// TIA Portal project "SortingStation" (V19)

(* hardware
DEVICE "S7-1500/ET200MP station_1"  S7-1500 station
   slot 0: "Rail_0"  Rack  6ES7 590-1***0-0AA0
   slot 1: "PLC_1"  CPU 1511-1 PN  6ES7 511-1AK02-0AB0  V2.9
      slot 3: "CPU display_1"  6ES7591-1AA00-0AA0
      slot 32768: "PROFINET interface_1"  X1
         slot 32769: "Port_1"  X1 P1
         slot 32770: "Port_2"  X1 P2
      slot 34817: "Virtual CP interface port_1"  Virtual CP interface port  Virtual CP interface port
   slot 2: "DI 16x24VDC BA_1"  DI 16x24VDC BA  6ES7 521-1BH10-0AA0  V1.1
   slot 3: "DQ 16x24VDC/0.5A BA_1"  DQ 16x24VDC/0.5A BA  6ES7 522-1BH10-0AA0  V1.1
   slot 4: "AI 4xU/I/RTD/TC ST_1"  AI 4xU/I/RTD/TC ST  6ES7 531-7QD00-0AB0  V1.0
DEVICE "HMI_1"  TP700 Comfort
   slot 0: "HMI_1"  TP700 Comfort  6AV2 124-0GC01-0AX0  17.0.0.0
   slot 1: "HMI_RT_1"  TP700 Comfort  6AV2 124-0GC01-0AX0  17.0.0.0
   slot 5: "HMI_1.IE_CP_1"  PROFINET Interface  17.0.0.0
      slot 1: "PROFINET Interface_1"  PROFINET Interface
         slot 1: "Port_1"  Port
         slot 2: "Port_2"  Port
   slot 7: "HMI_1.MPI/DP_CP_1"  MPI/DP Interface  17.0.0.0
*)

// ===== PLC "PLC_1"  CPU 1511-1 PN =====

VAR_GLOBAL   // PLC tag table "Default tag table"
   "System_Byte" AT %MB1 : Byte;
   "FirstScan" AT %M1.0 : Bool;
   "DiagStatusUpdate" AT %M1.1 : Bool;
   "AlwaysTRUE" AT %M1.2 : Bool;
   "AlwaysFALSE" AT %M1.3 : Bool;
   "Clock_Byte" AT %MB0 : Byte;
   "Clock_10Hz" AT %M0.0 : Bool;
   "Clock_5Hz" AT %M0.1 : Bool;
   "Clock_2.5Hz" AT %M0.2 : Bool;
   "Clock_2Hz" AT %M0.3 : Bool;
   "Clock_1.25Hz" AT %M0.4 : Bool;
   "Clock_1Hz" AT %M0.5 : Bool;
   "Clock_0.625Hz" AT %M0.6 : Bool;
   "Clock_0.5Hz" AT %M0.7 : Bool;
END_VAR

VAR_GLOBAL   // PLC tag table "IO_Tags"
   "PB_Start" AT %I0.0 : Bool;   // Start pushbutton, NO contact
   "PB_Stop" AT %I0.1 : Bool;   // Stop pushbutton, NC contact
   "PB_Reset" AT %I0.2 : Bool;   // Alarm reset pushbutton
   "ESTOP_OK" AT %I0.3 : Bool;   // Emergency stop circuit, 1 = healthy
   "S_Entry" AT %I0.4 : Bool;   // Part entry sensor
   "S_Defective" AT %I0.5 : Bool;   // Defective part signal
   "Motor_Overload_OK" AT %I0.6 : Bool;   // Motor overload relay, NC, 1 = healthy
   "AI_MotorTemp" AT %IW64 : Int;   // Motor temperature, raw analog value 0..27648
   "K_Motor" AT %Q0.0 : Bool;   // Conveyor motor contactor
   "L_Run" AT %Q0.1 : Bool;   // Green lamp, running
   "L_Fault" AT %Q0.2 : Bool;   // Red lamp, fault
   "L_Idle" AT %Q0.3 : Bool;   // Yellow lamp, idle
   "Y_Diverter" AT %Q0.4 : Bool;   // Diverter actuator for rejected parts
   "Horn" AT %Q0.5 : Bool;   // Alarm horn
END_VAR

TYPE "udt_Station"
   STRUCT
      State : Int;   // 0=Idle, 1=Running, 2=Fault
      FaultCode : Word := 0;   // bit0=EStop, bit1=Overload, bit2=OverTemp, bit3=Jam
      CntGood : DInt := 0;   // Count of good parts
      CntReject : DInt;   // Count of rejected parts
      MotorTemp : Real;   // Scaled motor temperature in degC
      TempLimit : Real := 80.0;   // Max allowed motor temperature in degC
      HMI_Start : Bool;   // Start command from HMI
      HMI_Stop : Bool;   // Stop command from HMI
      HMI_Reset : Bool;   // Alarm reset command from HMI
      HMI_ResetCnt : Bool;   // Counter reset command from HMI
   END_STRUCT;
END_TYPE

DATA_BLOCK "DB_Station"   // DB1
{ S7_Optimized_Access := 'TRUE' }
VERSION : 0.1
BEGIN
END_DATA_BLOCK

DATA_BLOCK "iDB_Station"   // DB2
{ S7_Optimized_Access := 'TRUE' }
VERSION : 0.1
// stored: InstanceOfName FB_Station
"FB_Station"
BEGIN
END_DATA_BLOCK

FUNCTION_BLOCK "FB_Motor"   // FB1, LAD
{ S7_Optimized_Access := 'TRUE' }
VERSION : 0.1
   VAR_INPUT
      Start : Bool;   // Start command, 1 = start requested
      Stop : Bool;   // Stop command, 1 = stop requested
      Permissive : Bool;   // Interlock, 1 = all conditions healthy
   END_VAR
   VAR_OUTPUT
      Run : Bool;   // Motor run command
   END_VAR
   VAR
      RunMem : Bool;   // Seal-in memory bit
   END_VAR
BEGIN

REGION Network 1: Seal-in memory bit
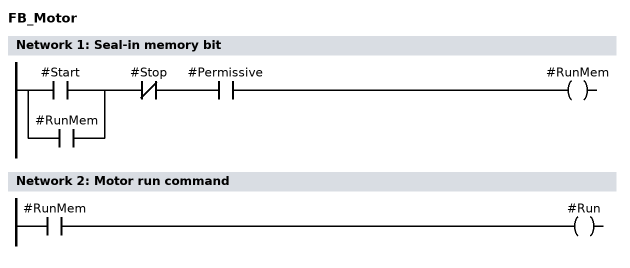
   RUNG wire#powerrail
      Contact( #Start )
      wire#w1
      I_Contact( #Stop )
      Contact( #Permissive )
      Coil( #RunMem )
   END_RUNG
   RUNG wire#powerrail
      Contact( #RunMem )
   END_RUNG wire#w1
   // the same network as SCL:
   #RunMem := (#Start OR #RunMem) AND NOT #Stop AND #Permissive;
END_REGION

REGION Network 2: Motor run command
   RUNG wire#powerrail
      Contact( #RunMem )
      Coil( #Run )
   END_RUNG
   // the same network as SCL:
   #Run := #RunMem;
END_REGION
END_FUNCTION_BLOCK

FUNCTION_BLOCK "FB_Station"   // FB2, SCL
{ S7_Optimized_Access := 'TRUE' }
VERSION : 0.1
   VAR_INPUT
      PB_Start : Bool;   // Start pushbutton, NO
      PB_Stop : Bool;   // Stop pushbutton, NC, 0 = pressed
      PB_Reset : Bool;   // Alarm reset pushbutton
      ESTOP_OK : Bool;   // Emergency stop circuit, 1 = healthy
      S_Entry : Bool;   // Part entry sensor
      S_Defective : Bool;   // Defective part signal
      Motor_Overload_OK : Bool;   // Overload relay, 1 = healthy
      Clock1Hz : Bool;   // 1 Hz clock bit for blinking
   END_VAR
   VAR_OUTPUT
      K_Motor : Bool;   // Conveyor motor contactor
      L_Run : Bool;   // Green lamp
      L_Fault : Bool;   // Red lamp, blinking
      L_Idle : Bool;   // Yellow lamp
      Y_Diverter : Bool;   // Diverter for rejected parts
      Horn : Bool;   // Alarm horn
   END_VAR
   VAR_IN_OUT
      Station : "udt_Station";   // Station data, passed from DB_Station
   END_VAR
   VAR
      motor : "FB_Motor";   // Motor control instance
      tonJam : TON_TIME;   // Jam detection timer
      tpDiverter : TP_TIME;   // Diverter pulse timer
   END_VAR
   VAR RETAIN
      ctuGood : CTU_DINT;   // Good parts counter
      ctuReject : CTU_DINT;   // Rejected parts counter
   END_VAR
   VAR
      rtStart : R_TRIG;   // Start edge
      rtReset : R_TRIG;   // Reset edge
      rtEntry : R_TRIG;   // Entry sensor edge
   END_VAR
   VAR_TEMP
      stopCmd : Bool;
      anyFault : Bool;
      fEStop : Bool;
      fOverload : Bool;
      fOverTemp : Bool;
      fJam : Bool;
      goodPulse : Bool;
      rejectPulse : Bool;
   END_VAR
BEGIN
   // =====================================================
   // FB_Station : sorting station main logic
   // States: 0 = Idle, 1 = Running, 2 = Fault
   // FaultCode: bit0 EStop, bit1 Overload, bit2 OverTemp, bit3 Jam
   // =====================================================

   // ---- 1. Edge detection and commands ----
   #rtStart(CLK := #PB_Start OR #Station.HMI_Start);
   #rtReset(CLK := #PB_Reset OR #Station.HMI_Reset);
   #rtEntry(CLK := #S_Entry);

   // PB_Stop is NC: 0 = pressed
   #stopCmd := (NOT #PB_Stop) OR #Station.HMI_Stop;

   // ---- 2. Fault detection (live conditions) ----
   #fEStop := NOT #ESTOP_OK;
   #fOverload := NOT #Motor_Overload_OK;
   #fOverTemp := #Station.MotorTemp > #Station.TempLimit;

   // Jam: entry sensor active longer than 5 s while running
   #tonJam(IN := #S_Entry AND (#Station.State = 1),
           PT := T#5s);
   #fJam := #tonJam.Q;

   #anyFault := #fEStop OR #fOverload OR #fOverTemp OR #fJam;

   // ---- 3. Latched fault code ----
   // Reset clears the code first, then active faults set their bits again
   IF #rtReset.Q THEN
       #Station.FaultCode := W#16#0000;
   END_IF;

   IF #fEStop THEN
       #Station.FaultCode := #Station.FaultCode OR W#16#0001;
   END_IF;
   IF #fOverload THEN
       #Station.FaultCode := #Station.FaultCode OR W#16#0002;
   END_IF;
   IF #fOverTemp THEN
       #Station.FaultCode := #Station.FaultCode OR W#16#0004;
   END_IF;
   IF #fJam THEN
       #Station.FaultCode := #Station.FaultCode OR W#16#0008;
   END_IF;

   // ---- 4. State machine ----
   CASE #Station.State OF
       0:  // Idle
           IF #anyFault THEN
               #Station.State := 2;
           ELSIF #rtStart.Q AND NOT #stopCmd THEN
               #Station.State := 1;
           END_IF;

       1:  // Running
           IF #anyFault THEN
               #Station.State := 2;
           ELSIF #stopCmd THEN
               #Station.State := 0;
           END_IF;

       2:  // Fault: leave only on reset with all faults cleared
           IF #rtReset.Q AND NOT #anyFault THEN
               #Station.State := 0;
           END_IF;

       ELSE
           #Station.State := 2;
   END_CASE;

   // ---- 5. Sorting logic (only while running) ----
   #goodPulse := FALSE;
   #rejectPulse := FALSE;

   IF (#Station.State = 1) AND #rtEntry.Q THEN
       IF #S_Defective THEN
           #rejectPulse := TRUE;
       ELSE
           #goodPulse := TRUE;
       END_IF;
   END_IF;

   #ctuGood(CU := #goodPulse,
            R := #Station.HMI_ResetCnt,
            PV := 99999999);
   #ctuReject(CU := #rejectPulse,
              R := #Station.HMI_ResetCnt,
              PV := 99999999);
   #Station.CntGood := #ctuGood.CV;
   #Station.CntReject := #ctuReject.CV;

   // Diverter: 2 s pulse for each rejected part
   #tpDiverter(IN := #rejectPulse,
               PT := T#2s);
   #Y_Diverter := #tpDiverter.Q AND (#Station.State = 1);

   // ---- 6. Motor control ----
   // Permissive drops the motor in Idle and Fault
   #motor(Start := #PB_Start OR #Station.HMI_Start,
          Stop := #stopCmd,
          Permissive := (#Station.State = 1));
   #K_Motor := #motor.Run;

   // ---- 7. Lamps and horn ----
   #L_Idle := (#Station.State = 0);
   #L_Run := (#Station.State = 1);
   #L_Fault := (#Station.State = 2) AND #Clock1Hz;
   #Horn := (#Station.State = 2);
END_FUNCTION_BLOCK

ORGANIZATION_BLOCK "Main"   // OB1, LAD, ProgramCycle
TITLE = "Main Program Sweep (Cycle)"
{ S7_Optimized_Access := 'TRUE' }
VERSION : 0.1
   VAR_INPUT
      Initial_Call : Bool;   // Initial call of this OB
      Remanence : Bool;   // =True, if remanent data are available
   END_VAR
   VAR_TEMP
      normTemp : Real;   // Normalized temperature 0.0 to 1.0
   END_VAR
BEGIN

REGION Network 1
   // Scale raw analog value 0..27648 to 0..150 degC
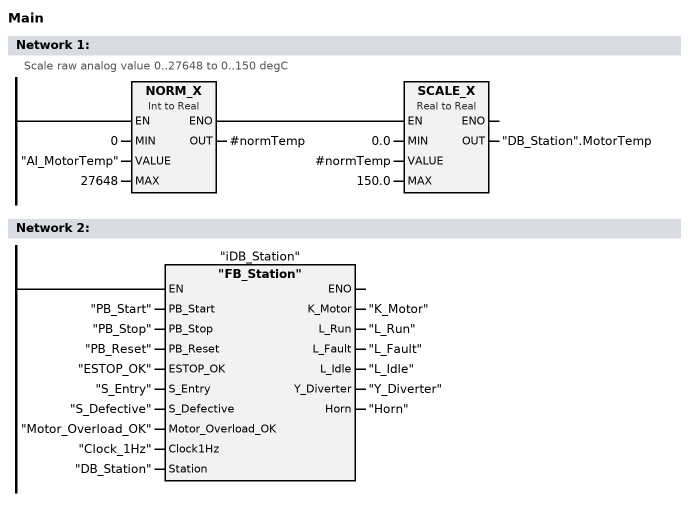
   RUNG wire#powerrail
      { S7_Templates := "[SrcType := Int, DestType := Real]" } Normalize(min := 0, value := "AI_MotorTemp", max := 27648, out => #normTemp)
      { S7_Templates := "[SrcType := Real, DestType := Real]" } Scale(min := 0.0, value := #normTemp, max := 150.0, out => "DB_Station".MotorTemp)
   END_RUNG
   // the same network as SCL:
   #normTemp := NORM_X(MIN := 0, VALUE := "AI_MotorTemp", MAX := 27648);
   "DB_Station".MotorTemp := SCALE_X(MIN := 0.0, VALUE := #normTemp, MAX := 150.0);
END_REGION

REGION Network 2
   RUNG wire#powerrail
      "iDB_Station"(PB_Start := "PB_Start", PB_Stop := "PB_Stop", PB_Reset := "PB_Reset", ESTOP_OK := "ESTOP_OK", S_Entry := "S_Entry", S_Defective := "S_Defective", Motor_Overload_OK := "Motor_Overload_OK", Clock1Hz := "Clock_1Hz", Station := "DB_Station", K_Motor => "K_Motor", L_Run => "L_Run", L_Fault => "L_Fault", L_Idle => "L_Idle", Y_Diverter => "Y_Diverter", Horn => "Horn")
   END_RUNG
   // the same network as SCL:
   "iDB_Station"(PB_Start := "PB_Start",   // "FB_Station"
                 PB_Stop := "PB_Stop",
                 PB_Reset := "PB_Reset",
                 ESTOP_OK := "ESTOP_OK",
                 S_Entry := "S_Entry",
                 S_Defective := "S_Defective",
                 Motor_Overload_OK := "Motor_Overload_OK",
                 Clock1Hz := "Clock_1Hz",
                 Station := "DB_Station",
                 K_Motor => "K_Motor",
                 L_Run => "L_Run",
                 L_Fault => "L_Fault",
                 L_Idle => "L_Idle",
                 Y_Diverter => "Y_Diverter",
                 Horn => "Horn");
END_REGION
END_ORGANIZATION_BLOCK

ORGANIZATION_BLOCK "Startup"   // OB100, SCL, Startup
TITLE = "Complete Restart"
{ S7_Optimized_Access := 'TRUE' }
VERSION : 0.1
   VAR_INPUT
      LostRetentive : Bool;   // True if retentive data are lost
      LostRTC : Bool;   // True if date and time are lost
   END_VAR
BEGIN
   // =====================================================
   // OB100 Startup : runs once at every STOP to RUN transition
   // Puts the station in a known safe state
   // =====================================================
   "DB_Station".State := 0;
   "DB_Station".FaultCode := W#16#0000;

   "DB_Station".HMI_Start := FALSE;
   "DB_Station".HMI_Stop := FALSE;
   "DB_Station".HMI_Reset := FALSE;
   "DB_Station".HMI_ResetCnt := FALSE;
END_ORGANIZATION_BLOCK

(* ===== HMI "HMI_RT_1" =====
system functions are stored by id; their names below are inferred from use
connection "HMI_Connection_1": ETHERNET, S7_1500_OMS

HMI tags "Default tag table"
   "Tag_ScreenNumber" : UInt, internal
   "Station_State" : Int = PLC DB_Station.State, 1 s
   "Station_FaultCode" : Word = PLC DB_Station.FaultCode AT %DB1.DBW0, 1 s
   "Station_CntGood" : DInt = PLC DB_Station.CntGood AT %DB1.DBW0, 1 s
   "Station_CntReject" : DInt = PLC DB_Station.CntReject AT %DB1.DBD0, 1 s
   "Station_MotorTemp" : Real = PLC DB_Station.MotorTemp AT %DB1.DBD0, 1 s
   "Station_TempLimit" : Real = PLC DB_Station.TempLimit AT %DB1.DBD0, 1 s
   "Station_HMI_Start" : Bool = PLC DB_Station.HMI_Start AT %DB1.DBD0, 1 s
   "Station_HMI_Stop" : Bool = PLC DB_Station.HMI_Stop AT %DB1.DBX0.0, 1 s
   "Station_HMI_Reset" : Bool = PLC DB_Station.HMI_Reset AT %DB1.DBX0.0, 1 s
   "Station_HMI_ResetCnt" : Bool = PLC DB_Station.HMI_ResetCnt AT %DB1.DBX0.0, 1 s

screen "Root screen" 800x420, template "Template_1"
   on GenerateScreen: SetTag("Tag_ScreenNumber", 1)
   TextField "HmiScreenItemData" at 78,377 size 640x25; Text 'Welcome to HMI_1 (TP700 Comfort)!'
   TextField "Text field_1" at 31,11 size 209x34; Text 'Sorting Station'
   TextField "Text field_2" at 78,70 size 54x23; Text 'State'
   TextField "Text field_3" at 77,113 size 51x23; Text 'Good'
   TextField "Text field_4" at 54,157 size 86x23; Text 'Rejected'
   TextField "Text field_5" at 19,201 size 123x23; Text 'Temperature'
   TextField "Text field_6" at 43,247 size 99x23; Text 'Fault code'
   IOField "I/O field_1" at 142,67 size 96x32; FormatPattern 9
      ProcessValue <- "Station_State"
   IOField "I/O field_2" at 142,108 size 96x32; FormatPattern 99999
      ProcessValue <- "Station_CntGood"
   IOField "I/O field_3" at 143,152 size 96x32; FormatPattern 99999
      ProcessValue <- "Station_CntReject"
   IOField "I/O field_4" at 143,197 size 96x32; FormatPattern 999.9
      ProcessValue <- "Station_MotorTemp"
   IOField "I/O field_5" at 143,246 size 96x32; FormatPattern FFFF
      ProcessValue <- "Station_FaultCode"
   Button "Button_1" at 384,75 size 96x32; TextOff 'Start'
      on Press: SetBit("Station_HMI_Start")
      on Release: ResetBit("Station_HMI_Start")
   Button "Button_2" at 383,128 size 96x32; TextOff 'Stop'
      on Press: SetBit("Station_HMI_Stop")
      on Release: ResetBit("Station_HMI_Stop")
   Button "Button_3" at 384,184 size 96x32; TextOff 'Reset'
      on Press: SetBit("Station_HMI_Reset")
      on Release: ResetBit("Station_HMI_Reset")
   Button "Button_4" at 384,238 size 141x32; TextOff 'Reset counters'
      on Press: SetBit("Station_HMI_ResetCnt")
      on Release: ResetBit("Station_HMI_ResetCnt")
   Circle "Circle_1" at 598,133 size 80x80
      Appearance <- "Station_State"
   TextField "Text field_8" at 239,201 size 50x23; Text 'degC'
*)